(* CODESYS project ROTATOR.project
   CustomField04_name: CustomField04
   CustomField06_name: CustomField06
   CustomField07_name: CustomField07
   CustomField09_name: CustomField09
   CustomField08_name: CustomField08
   CustomField02_name: CustomField02
   CustomField10_name: CustomField10
   CustomField01_name: CustomField01
   CustomField03_name: CustomField03
   CustomField05_name: CustomField05

Project tree, tasks and I/O mapping:
  Cebora : TM241CEC24T/U, Schneider Electric, order no. TM241CEC24T/U, version 4.0.6.18
      settings: OPCUA enable = False
    application Application
      libraries: Toolbox, 2.2.0.0 (Schneider Electric)
      task MAST (cyclic, interval 20 ms, priority 15, watchdog 100 ms x 1) calls Main
      global variables GVL
      program SndRecvRS232 [CFC]
      program Data_transfer [ST]
      program Motor [ST]
      program Main [ST]
      trace Trace (task MAST): RS232Read
      trace Trace_1 (task MAST): 
      trace Trace_2 (task MAST): SM1_STOP
      trace Trace_3 (task MAST): RS232Read
      trace Trace_4 (task ): , RS232Read
    Ethernet_1 : Ethernet Network, Schneider Electric, version 4.0.6.18
    COM_Bus : COM bus, Schneider Electric, version 4.0.6.18
    Counters : Counters, Schneider Electric, version 4.0.6.18
    IO_Bus : IO bus - TM3, Schneider Electric, version 4.0.6.18
    Serial_Line_1 : Serial line, Schneider Electric, version 4.0.6.18
      ROBOT : ASCII Manager, Schneider Electric, version 4.0.0.2
    Cartridge_1 : Cartridge, Schneider Electric, version 4.0.6.18
    Pulse_Generators : Pulse Generators, Schneider Electric, version 4.0.6.18
        settings: Instance name = 'SM1'; B output History = 'old=-1 new=1'; A output History = 'old=-1 new=0'; Temporary Instance name = 'SM1'
    DQ : Digital Outputs, Schneider Electric, version 4.0.6.18
        settings: Outputs Usage = 3
        unmapped channels: QW0, QB1
    CAN_1 : CANopen bus, Schneider Electric, version 4.0.6.18
    IO : Digital Inputs, Schneider Electric, version 4.0.6.18
        unmapped channels: IW0, IB1
    Serial_Line_2 : Serial line, Schneider Electric, version 4.0.6.18
*)

// Cebora/Application/GVL
VAR_GLOBAL	
	RS232_READ: SEND_RECV_MSG;
	RS232_SEND: SEND_RECV_MSG;
	IX0_0 AT %IX0.0: BOOL;
	DI_LEFT AT %IX0.1: BOOL;
	DI_RIGHT AT %IX0.2: BOOL;
	DI_RESET AT %IX0.3: BOOL;
	ROTATOR_ACTIVE AT %QX0.4: BOOL;
	InArr:ARRAY [1..18] OF BYTE;
	InSET_Pose:ARRAY [1..255] OF BYTE;
	InSET_Speed:ARRAY [1..255] OF BYTE;
	InStrSET_Pose:STRING;
	InStrSET_Speed:STRING;
	InRealSET_Pose:REAL;
	InRealSET_Speed:REAL;
	InBoolSET_Move: BOOL;
	
	RealGET_Pose: REAL;
	StrGET_Pose: STRING;
	OutArr:ARRAY [1..11] OF BYTE;	
	ArrGET_Pose:ARRAY [1..255] OF BYTE;
	
	RS232Read:BOOL;
	RS232Send:BOOL;
	Readed:BOOL;
	Sended:BOOL;
	T0:TON;
	T0_STATE:BOOL;
	T1:TON;
	T1_STATE:BOOL;
	T2:TON;
	T2_STATE:BOOL;
	T3:TON;
	T3_STATE:BOOL;
	T4:TON;
	T4_ActTime:TIME;
	//STOP_Read:BOOL;
	//StopReadTrig:BOOL;
	
	MC_Power_SM1: MC_Power_PTO;
	MC_Home_SM1: MC_Home_PTO;
	MC_MoveVelocity_SM1: MC_MoveVelocity_PTO;
	MC_Stop_SM1: MC_Stop_PTO;
	MC_MoveAbsolute_SM1: MC_MoveAbsolute_PTO;
	MC_MoveRelative_SM1: MC_MoveRelative_PTO;
	MC_ReadActualPosition_SM1: MC_ReadActualPosition_PTO;
	MC_SetPosition_SM1: MC_SetPosition_PTO;	
	SM1_RESOLUTION: REAL; //Кількість імп. на оберт
	SM1_SET_SPEED: REAL; //Фактичне задання швидкості
	SM1_SET_POSE: REAL; //Фактичне задання швидкості
	SM1_SET_MOVE: BOOL; //Фактичне значення старту
	Previous_SET_Pose: REAL; //Відслідковування зміни в позиції
	Previous_SET_Speed: REAL; //Відслідковування зміни в швидкості
	SM1_SET_DIR: MC_DIRECTION; //Фактичне задання напрямку
	SourceGET_Pose: REAL; //Значення MC_ReadActualPosition_SM1
	SM1_ABSOLUTE_START: BOOL; //Старт SM1 в автоматичному режимі
	SM1_STOP: BOOL; //Стоп руху
	RESET_POSE: BOOL; //Ресет позиції
END_VAR

VAR_GLOBAL RETAIN
	
END_VAR

// Cebora/Application/Main
PROGRAM Main
VAR
END_VAR

SM1_RESOLUTION:= 100; //Кількість імпульсів на градус
Data_transfer();
Motor();

END_PROGRAM

// Cebora/Application/Data_transfer
PROGRAM Data_transfer

VAR
	I: INT;
	FB_6: SE_TBX.FB_Scaling;
	FB_5: SE_TBX.FB_Scaling;
	FB_4: SE_TBX.FB_Scaling;
	FB_3: SE_TBX.FB_Scaling;
	FB_2: SE_TBX.FB_Scaling;
	FB_1: SE_TBX.FB_Scaling;
	FB_0: SE_TBX.FB_Scaling;;
END_VAR

	RS232Send:= FALSE;
	RS232Read:= TRUE; 
	SndRecvRS232(); 
	RS232Read:= FALSE; 
	SndRecvRS232();

		//Reading data
		IF 	InArr[1] = 83 AND InArr[18] = 70 THEN //Умова задання даних
			FOR I:= 1 TO 9 BY 1 DO
				InSET_Pose[I]:= InArr[I+1];
			END_FOR
			FOR I:= 1 TO 6 BY 1 DO
				InSET_Speed[I]:= InArr[I+10];
			END_FOR
			InStrSET_Pose:= ArrayOfByte_TO_String(i_abyIput:= InSET_Pose, i_xOrdr:= TRUE , i_xSpce:=  FALSE);
			InStrSET_Speed:= ArrayOfByte_TO_String(i_abyIput:= InSET_Speed, i_xOrdr:= TRUE , i_xSpce:=  FALSE);
			InRealSET_Pose:= STRING_TO_REAL(InStrSET_Pose); //Set Pose
			InRealSET_Speed:= STRING_TO_REAL(InStrSET_Speed); //Set Speed
			IF InArr[17] = 49 THEN InBoolSET_Move:= TRUE; ELSE InBoolSET_Move:= FALSE; END_IF 
		END_IF
		//Reading data
		
		IF RESET_POSE THEN InArr[17]:= 48; InBoolSET_Move:= FALSE; END_IF //Reset move from button
		
		//Reset speed from button
		IF RESET_POSE THEN 
			FOR I:= 1 TO 6 BY 1 DO
				InArr[11]:= 48; InArr[12]:= 49; InArr[13]:= 48; InArr[14]:= 46; InArr[15]:= 48; InArr[16]:= 48;
				InSET_Speed[I]:= InArr[I+10];
			END_FOR
			InStrSET_Speed:= ArrayOfByte_TO_String(i_abyIput:= InSET_Speed, i_xOrdr:= TRUE , i_xSpce:=  FALSE);
			InRealSET_Speed:= STRING_TO_REAL(InStrSET_Speed); //Set Speed
		END_IF
		//Reset speed from button
		
		//Sending data calculation
		OutArr[1]:= 83;
		RealGET_Pose:= SourceGET_Pose / SM1_RESOLUTION;
		StrGET_Pose:= REAL_TO_STRING(RealGET_Pose);
		ArrGET_Pose:= String_TO_ArrayOfByte(i_sIput:= StrGET_Pose,i_xOrdr:= TRUE);
		FOR I:= 1 TO 9 BY 1 DO
			OutArr[I+1]:= ArrGET_Pose[I];
			IF OutArr[I+1] = 0 THEN OutArr[I+1]:= 48; END_IF
		END_FOR;
		OutArr[11]:= 70;
		//Sending data calculation
		
		//Sending data
		IF InArr[1] = 82 AND InArr[18] = 80 THEN //Умова відправки даних (поточна позиція)
			RS232Read:= FALSE;
			RS232Send:= TRUE;
			SndRecvRS232();
			RS232Send:= FALSE;
			SndRecvRS232();
		END_IF
		//Sending data

END_PROGRAM

// Cebora/Application/SndRecvRS232
PROGRAM SndRecvRS232
VAR
	ADDM1: ADDM;
	ADDM2: ADDM;
	myAddressTable: ADDRESS;
END_VAR

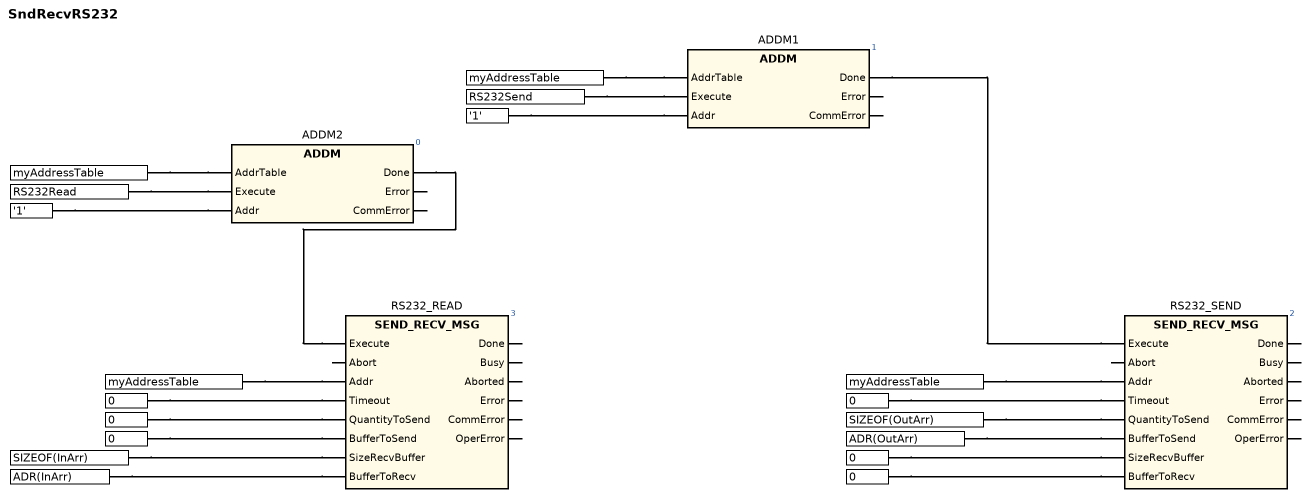
ADDM2(AddrTable := myAddressTable, Execute := RS232Read, Addr := '1'); // ADDM
ADDM1(AddrTable := myAddressTable, Execute := RS232Send, Addr := '1'); // ADDM
RS232_SEND(
    Execute := ADDM1.Done,
    Addr := myAddressTable,
    Timeout := 0,
    QuantityToSend := SIZEOF(OutArr),
    BufferToSend := ADR(OutArr),
    SizeRecvBuffer := 0,
    BufferToRecv := 0); // SEND_RECV_MSG
RS232_READ(
    Execute := ADDM2.Done,
    Addr := myAddressTable,
    Timeout := 0,
    QuantityToSend := 0,
    BufferToSend := 0,
    SizeRecvBuffer := SIZEOF(InArr),
    BufferToRecv := ADR(InArr)); // SEND_RECV_MSG

END_PROGRAM

// Cebora/Application/Motor
PROGRAM Motor
VAR
	RESET_POSE_TON: TON;
	MC_POWER_DELAY: TON;
	INIT_TRIG: BOOL;
	SM1_START_TRIG: F_TRIG;
	SM1_STOP_RIGHT: F_TRIG;
	SM1_STOP_AUTO: F_TRIG;
	SM1_STOP_LEFT: F_TRIG;
	T1_START: TON;
	SET_MOVE_TRIG: R_TRIG;
	FIRST_MOTOR_ENA: R_TRIG;
	FIRST_MOTOR_ENA_DONE: BOOL;
	TON_RESET_POS: TON;
	SM1_DIRECTION: MC_DIRECTION;
	FIRST_START: BOOL ;
END_VAR

MC_POWER_DELAY(IN:=NOT INIT_TRIG , PT:=T#100MS , Q=> , ET=> ); //Затримка ініціалізації
IF MC_POWER_DELAY.Q THEN INIT_TRIG:=TRUE; END_IF; //Затримка ініціалізації
IF MC_POWER_SM1.Error THEN INIT_TRIG:=FALSE; END_IF; //Ресет при виникненні помилки

IF (NOT FIRST_START AND INIT_TRIG) OR DI_RESET THEN FIRST_START:= TRUE; RESET_POSE:= TRUE; END_IF //Ресет позиції
RESET_POSE_TON(IN:=RESET_POSE , PT:=T#100MS); //Затримка на скидання тригеру ресету позиції
IF RESET_POSE_TON.Q THEN RESET_POSE:= FALSE; END_IF //Скидання тригеру ресету позиції

SM1_SET_POSE:= InRealSET_Pose; //Задання позиції
IF (DI_LEFT OR DI_RIGHT) AND InRealSET_Speed = 0 THEN SM1_SET_SPEED:= 10; ELSE SM1_SET_SPEED:= InRealSET_Speed; END_IF //Логіка задання швидкості
IF DI_LEFT THEN SM1_SET_DIR:= -1; ELSIF DI_RIGHT THEN SM1_SET_DIR:= 1; END_IF //Логіка задання напрямку

SM1_SET_MOVE:= InBoolSET_Move; //Задання старту/стопу
SET_MOVE_TRIG(CLK:= InBoolSET_Move); //Для старту після зупинки, якщо не змінювалась швидкість і позиція
IF ((SM1_SET_POSE <> Previous_SET_Pose OR SM1_SET_SPEED <> Previous_SET_Speed) AND NOT (DI_LEFT OR DI_RIGHT) AND SM1_SET_MOVE) OR SET_MOVE_TRIG.Q THEN //Старт автомат
SM1_ABSOLUTE_START:= TRUE; Previous_SET_Pose:= SM1_SET_POSE; Previous_SET_Speed:= SM1_SET_SPEED; ELSE SM1_ABSOLUTE_START:= FALSE; END_IF //Старт автомат

SM1_STOP_LEFT(CLK:= DI_LEFT); //Тригер стопу в ручному режимі
SM1_STOP_RIGHT(CLK:= DI_RIGHT); //Тригер стопу в ручному режимі
SM1_STOP_AUTO(CLK:= InBoolSET_Move); //Тригер стопу в автоматичному режимі
IF SM1_STOP_LEFT.Q OR SM1_STOP_RIGHT.Q OR SM1_STOP_AUTO.Q THEN SM1_STOP:= TRUE; END_IF //Стоп руху автомат по тригеру
IF MC_Stop_SM1.Done THEN SM1_STOP:=  FALSE; END_IF //Стоп руху

MC_Power_SM1(
	Axis:=SM1 , 
	Enable:=INIT_TRIG , 
	DriveReady:=TRUE , 
	LimP:=TRUE , 
	LimN:=TRUE , 
	Status=> , 
	DriveEnable=> , 
	Error=> , 
	ErrorId=> );

//РУХ В АВТОМАТІ ПО АБСОЛЮТНИХ ПОЗИЦІЯХ	
MC_MoveAbsolute_SM1(
	Axis:=SM1 , 
	Execute:= SM1_ABSOLUTE_START, 
	Position:= REAL_TO_DINT(SM1_SET_POSE * SM1_RESOLUTION), 
	Velocity:= REAL_TO_DINT(SM1_SET_SPEED * SM1_RESOLUTION), 
	Acceleration:= 200, 
	Deceleration:= 200, 
	BufferMode:= , 
	Done=> , 
	Busy=> , 
	Active=> , 
	CommandAborted=> , 
	Error=> , 
	ErrorId=> , 
	JerkRatio:= );
//РУХ В АВТОМАТІ ПО АБСОЛЮТНИХ ПОЗИЦІЯХ	

IF NOT MC_MoveAbsolute_SM1.Busy AND NOT MC_MoveAbsolute_SM1.Active THEN ROTATOR_ACTIVE:=FALSE; ELSE ROTATOR_ACTIVE:=TRUE; END_IF //Фізичний вихід для слідкування зайнятості двигуна

//РУХ В РУЧНОМУ
MC_MoveVelocity_SM1(
	Axis:=SM1 , 
	Execute:= (DI_LEFT OR DI_RIGHT) AND NOT ROTATOR_ACTIVE, 
	ContinuousUpdate:= TRUE, 
	Velocity:= REAL_TO_DINT(SM1_SET_SPEED * SM1_RESOLUTION),
	Acceleration:= 200, 
	Deceleration:= 200, 
	Direction:= SM1_SET_DIR, 
	BufferMode:= , 
	InVelocity=> , 
	Busy=> , 
	Active=> , 
	CommandAborted=> , 
	Error=> , 
	ErrorId=> , 
	JerkRatio:= );
//РУХ В РУЧНОМУ
	
MC_ReadActualPosition_SM1(
	Axis:=SM1 , 
	Enable:=TRUE , 
	Valid=> , 
	Error=> , 
	ErrorId=> ,
	Position=> );
	
SourceGET_Pose:= DINT_TO_REAL(MC_ReadActualPosition_SM1.Position); //Читання поточної позиції

MC_SetPosition_SM1(
	Axis:=SM1 , 
	Execute:= RESET_POSE,
	Position:= 0, 
	Done=> , 
	Error=> , 
	ErrorId=> );
	
MC_Stop_SM1(
	Axis:=SM1 , 
	Execute:= SM1_STOP,
	Deceleration:= , 
	Done=>, 
	Busy=> , 
	CommandAborted=> , 
	Error=> , 
	ErrorId=> , 
	JerkRatio:= );
	
{MC_Home_SM1(
	Axis:=SM1 , 
	Execute:= , 
	Mode:= , 
	Position:= , 
	Direction:= , 
	HighVelocity:= , 
	LowVelocity:= , 
	Acceleration:= , 
	Deceleration:= , 
	Offset:= , 
	Done=> , 
	Busy=> , 
	Active=> , 
	CommandAborted=> , 
	Error=> , 
	ErrorId=> , 
	JerkRatio:= );
	
MC_MoveRelative_SM1(
	Axis:=SM1 , 
	Execute:= , 
	Distance:= ,
	Velocity:= ,
	Acceleration:= , 
	Deceleration:= , 
	BufferMode:= , 
	Done=> , 
	Busy=> , 
	Active=> , 
	CommandAborted=> , 
	Error=> , 
	ErrorId=> , 
	JerkRatio:= );}

END_PROGRAM
